// TwinCAT 3 PLC project PLC1
// ProgramVersion: 3.1.4026.17
// libraries:
//   Tc2_Standard, * (Beckhoff Automation GmbH)
//   Tc2_System, * (Beckhoff Automation GmbH)
// project tree:
//   / PlcTask.TcTTO
//   POUs/ MAIN.TcPOU
// real-time tasks:
//   TASK PlcTask: cycle T#10ms, priority 20, ADS port 350

CONFIGURATION PLC1
    RESOURCE PLC ON TwinCAT3
        TASK PlcTask(INTERVAL := T#10ms, PRIORITY := 20);
        PROGRAM MAIN WITH PlcTask : MAIN;
    END_RESOURCE
END_CONFIGURATION

// ---- POUs/MAIN.TcPOU
PROGRAM MAIN
VAR
	Nivel1 		: INT := 0;
	Nivel1Cheio	: BOOL;
	Nivel2 		: INT := 0;
	BombaAtiva 	: BOOL;
	Timer		: TON;
END_VAR

IF NOT BombaAtiva AND Nivel1 < 100 THEN
	Nivel1 := Nivel1 + 1;
	IF Nivel1 = 100 THEN
		Nivel1 := 100;
		Nivel1Cheio := TRUE;
	END_IF
END_IF

Timer(IN:= Nivel1Cheio, PT:= T#5S, Q=> BombaAtiva);

IF BombaAtiva AND Nivel1 >= 100 THEN
	Nivel2 := Nivel2 + 1;
	IF Nivel2 = 100 THEN
		Nivel2 := 100;
		BombaAtiva := FALSE;
	END_IF
END_IF

END_PROGRAM
